// TIA Portal V21 export
// export: Created 2026-08-21T20:18:52.4212526Z, ExportSetting None, DisplayName Totally Integrated Automation Portal, DisplayVersion V21, DisplayName STEP 7 Professional, DisplayVersion V21, DisplayName STEP 7 Safety, DisplayVersion V21, DisplayName Tech WebApplication, DisplayVersion V21, DisplayName WinCC Basic/Comfort/Advanced, DisplayVersion V21, DisplayName WinCC Professional, DisplayVersion V21, DisplayName WinCC Unified, DisplayVersion V21
DATA_BLOCK "ServiceCommandLogicDB"   // DB11
// stored: InstanceOfName Service_Command_Logic, InstanceOfType FB
"Service_Command_Logic"
   // VAR_INPUT
   //    Level : Real;
   //    ProcedureID_cur : DWord;
   // END_VAR
BEGIN
END_DATA_BLOCK
